# EPICS autosave request: roles/device_roles/adphantom/files/auto_settings.req
file "ADBase_settings.req",          P=$(P),  R=cam1:
file "NDStdArrays_settings.req",    P=$(P),  R=image1:
file "commonPlugin_settings.req",   P=$(P)
